(* IEC 61131-3 sources: SortJet_MasterSPS_Aufbau.fbsproj/08_POUs/Basis Programmbausteine, 6 files *)

(* ---- AutomatischeFachaufnahme.prg.st ---- *)
(* METADATA
{
	"v3Meta": {
		"objectGuid": "2dd67d59-9d65-422a-a9a5-a54784296135"
	}
}
*)
PROGRAM AutomatischeFachaufnahme
VAR_INPUT

  // BOOLEAN
  bpStarteFachaufnahme : BOOL := FALSE;
  bpAktiv              : BOOL := TRUE;

  // WORD
  wpMMINummer  : WORD;

  // POINTER
  ptQuerfahrtShuttle : REFERENCE TO Rexroth_ctrlX_Drive_Eckelmann_MC_V01_02_02;

  // REF
  Shuttle : REFERENCE TO Shuttle_FB_V01_00_00;

END_VAR

VAR

  // STEP
  steplAufnahme            : STEPS_TE;

  // WORD

  // REAL
  rlLetztePosition         : REAL;
  rlMerkerGeschwindigkeit  : real;

  // POINTER
  ptlAnalogwertChannel1  : REFERENCE TO INT;
  ptlAnalogwertChannel2  : REFERENCE TO INT;

END_VAR

VAR CONSTANT

  // WORD
  wGeschwindigkeitFachaufnahme : WORD := 5;
  wDefaultHandgeschwindigkeit  : WORD := 300;

END_VAR

//-------------------------------------------------------------------------------------------------
// AUTOMATISIERTE FACHAUFNAHME
//-------------------------------------------------------------------------------------------------
(* Anmerkung:
   - Shuttle-Koordinationsbaustein zur Fachaufnahme
*)
IF ( bpAktiv ) THEN

  (* Hinweis:
     - Starten der Fachaufnahme
  *)
  Shuttle REF= aShuttle[wpMMINummer];
  IF NOT __ISVALIDREF(Shuttle) THEN
    RETURN;
  ELSE
    ptQuerfahrtShuttle    REF= Shuttle.Querfahrt.Antrieb;
    ptlAnalogwertChannel1 REF= Shuttle.in_iAnalogwertChannel1;
    ptlAnalogwertChannel2 REF= Shuttle.in_iAnalogwertChannel2;
  END_IF

  (* Hinweis:
     - Starten der Fachaufnahme
  *)
  IF ( bpStarteFachaufnahme ) THEN

    IF ( __ISVALIDREF(ptQuerfahrtShuttle) ) THEN

      CASE steplAufnahme OF

        // -----------------------------------------------------------------------
        STEP_0_E:
          rlMerkerGeschwindigkeit :=  ptQuerfahrtShuttle.ppAntriebsInformationen.rpHandGeschwindigkeit;
          ptQuerfahrtShuttle.ppAntriebsInformationen.rpHandGeschwindigkeit := wGeschwindigkeitFachaufnahme;

          steplAufnahme:= STEP_10_E;

        // -----------------------------------------------------------------------
        STEP_10_E:
          IF (  ( ptQuerfahrtShuttle.rpIstPosition <> rlLetztePosition )
               AND ( ptQuerfahrtShuttle.rpIstPosition <> 0 ) )
          THEN

            rlLetztePosition := ptQuerfahrtShuttle.rpIstPosition;

            (* Hinweis:
               - Nachricht an das HMI
            *)
            rSPS2MMIFachaufnahmePosition   := rlLetztePosition;
            wSPS2MMIFachaufnahmeAnalogwert := TO_WORD(ptlAnalogwertChannel1);
            MsgToMmi( SB0_SPS_FACHAUFNAHMEDATEN );
          END_IF

      END_CASE

    ELSE
      ;

    END_IF

  END_IF

  IF ( NOT bpStarteFachaufnahme ) THEN

    IF ( steplAufnahme > STEP_0_E ) THEN
      steplAufnahme := STEP_0_E;
      ptQuerfahrtShuttle.ppAntriebsInformationen.rpHandGeschwindigkeit := SEL( rlMerkerGeschwindigkeit <> 0, wDefaultHandgeschwindigkeit, rlMerkerGeschwindigkeit ) ;
      rlMerkerGeschwindigkeit := 0;
    END_IF

  END_IF

END_IF
END_PROGRAM

(* ---- CheckReset.prg.st ---- *)
(* METADATA
{
	"v3Meta": {
		"objectGuid": "ed448837-b746-4b1a-b2e7-236797e04e0f"
	}
}
*)
PROGRAM CheckReset
VAR
  wlIndexAutomatikkreis,
  wlIndexStation : WORD;
END_VAR

FOR wlIndexAutomatikkreis := cERSTER_AUTOMATIKKREIS TO cLETZTER_AUTOMATIKKREIS DO

  agbResetAktiv[wlIndexAutomatikkreis] := FALSE;

  FOR wlIndexStation := cERSTE_STATION TO cLETZTE_STATION DO
    IF starrStationBasisParameter[wlIndexStation].bReset AND_THEN StationInAutomatikkreis(starrStationBasisParameter[wlIndexStation].stMKs.eaAutomatikkreis, wlIndexAutomatikkreis) THEN
      agbResetAktiv[wlIndexAutomatikkreis] := TRUE;
      EXIT;
    END_IF
  END_FOR

  // Schleife des AK eine Iteration weiter
  IF agbResetAktiv[wlIndexAutomatikkreis] THEN
    CONTINUE;
  END_IF

  FOR wlIndexStation := cERSTES_SHUTTLE TO cLETZTES_SHUTTLE DO
    IF starrShuttleBasisParameter[wlIndexStation].bReset AND_THEN StationInAutomatikkreis(starrShuttleBasisParameter[wlIndexStation].stMKs.eaAutomatikkreis, wlIndexAutomatikkreis) THEN
      agbResetAktiv[wlIndexAutomatikkreis] := TRUE;
      EXIT;
    END_IF
  END_FOR

  // Schleife des AK eine Iteration weiter
  IF agbResetAktiv[wlIndexAutomatikkreis] THEN
    CONTINUE;
  END_IF

  FOR wlIndexStation := cERSTES_TRANSFERSHUTTLE TO cLETZTES_TRANSFERSHUTTLE DO
    IF starrTransferShuttleBasisParameter[wlIndexStation].bReset AND_THEN StationInAutomatikkreis(starrTransferShuttleBasisParameter[wlIndexStation].stMKs.eaAutomatikkreis, wlIndexAutomatikkreis) THEN
      agbResetAktiv[wlIndexAutomatikkreis] := TRUE;
      EXIT;
    END_IF
  END_FOR

  // Schleife des AK eine Iteration weiter
  IF agbResetAktiv[wlIndexAutomatikkreis] THEN
    CONTINUE;
  END_IF

  FOR wlIndexStation := cERSTE_FAECHERWAGENSTATIONS_NR TO cLETZTE_FAECHERWAGENSTATIONS_NR DO
    IF starrFaecherwagenBasisParameter[wlIndexStation].bReset AND_THEN StationInAutomatikkreis(starrFaecherwagenBasisParameter[wlIndexStation].stMKs.eaAutomatikkreis, wlIndexAutomatikkreis) THEN
      agbResetAktiv[wlIndexAutomatikkreis] := TRUE;
      EXIT;
    END_IF
  END_FOR

  // Schleife des AK eine Iteration weiter
  IF agbResetAktiv[wlIndexAutomatikkreis] THEN
    CONTINUE;
  END_IF

  FOR wlIndexStation := cERSTE_FREMDANLAGE_EINLAUF TO cLETZTE_FREMDANLAGE_EINLAUF DO
    IF starrFremdanlageEinlaufStationBasisParameter[wlIndexStation].bReset AND_THEN StationInAutomatikkreis(starrFremdanlageEinlaufStationBasisParameter[wlIndexStation].stMKs.eaAutomatikkreis, wlIndexAutomatikkreis) THEN
      agbResetAktiv[wlIndexAutomatikkreis] := TRUE;
      EXIT;
    END_IF
  END_FOR

  // Schleife des AK eine Iteration weiter
  IF agbResetAktiv[wlIndexAutomatikkreis] THEN
    CONTINUE;
  END_IF

  FOR wlIndexStation := cERSTE_FREMDANLAGE_AUSLAUF TO cLETZTE_FREMDANLAGE_AUSLAUF DO
    IF starrFremdanlageAuslaufStationBasisParameter[wlIndexStation].bReset AND_THEN StationInAutomatikkreis(starrFremdanlageAuslaufStationBasisParameter[wlIndexStation].stMKs.eaAutomatikkreis, wlIndexAutomatikkreis) THEN
      agbResetAktiv[wlIndexAutomatikkreis] := TRUE;
      EXIT;
    END_IF
  END_FOR

END_FOR
END_PROGRAM

(* ---- ErsteUndLetzteScheibeBits.prg.st ---- *)
(* METADATA
{
	"v3Meta": {
		"objectGuid": "2dfa9b46-65fe-42f1-b72f-b251bddaa00a"
	}
}
*)
PROGRAM ErsteUndLetzteScheibeBits
VAR_INPUT

  // WORD
  wpErsteUndLetzteScheibe : WORD;

END_VAR
VAR_OUTPUT

  // WORD
  wpLetzteScheibe,
  wpErsteScheibe   : WORD;

END_VAR
VAR

  // WORD
  wlMerkerErsteUndLetzteScheibe  : WORD;

END_VAR
VAR CONSTANT

  // WORD
  cBIT_MASKE_LETZTE_SCHEIBE  : WORD := 2#0000000011111111;

END_VAR

//-------------------------------------------------------------------------------------------------
// BAUSTEIN: LOGIK
//-------------------------------------------------------------------------------------------------

(* Hinweis:
   - Erste Scheibe
*)
wlMerkerErsteUndLetzteScheibe := wpErsteUndLetzteScheibe;
wpLetzteScheibe := wlMerkerErsteUndLetzteScheibe AND cBIT_MASKE_LETZTE_SCHEIBE;

(* Hinweis:
   - Letzte Scheibe
*)
wlMerkerErsteUndLetzteScheibe := wpErsteUndLetzteScheibe;
wpErsteScheibe := SHR(wlMerkerErsteUndLetzteScheibe, 8);
END_PROGRAM

(* ---- Schrittketten_Logger.prg.st ---- *)
(* METADATA
{
	"v3Meta": {
		"objectGuid": "cb3b1eb5-1dc3-4d16-abd2-ade96f8e42d9"
	}
}
*)
PROGRAM Schrittketten_Logger
VAR

  // WORD
  i              : WORD;
  j              : WORD;
  wiSchrittkette : ARRAY[0..7] OF WORD;
  wlSchrittkette : ARRAY[0..7,0..31] OF WORD;

  // STRING
  sBezeichnung   : ARRAY[0..7] OF STRING;

END_VAR
sBezeichnung[0]   := ' - ';
wiSchrittkette[0] := 0;

sBezeichnung[1]   := ' - ';
wiSchrittkette[1] := 0;

sBezeichnung[2]   :=  ' - ';
wiSchrittkette[2] :=  0;

sBezeichnung[3]   :=  ' - ';
wiSchrittkette[3] :=  0;

sBezeichnung[4]   := ' - ';
wiSchrittkette[4] := 0;

sBezeichnung[5]   := ' - ';
wiSchrittkette[5] := 0;

sBezeichnung[6]   := ' - ';
wiSchrittkette[6] := 0;

sBezeichnung[7]   := ' - ';
wiSchrittkette[7] := 0;

FOR i := 0 TO 7 DO

  IF(wiSchrittkette[i] <> wlSchrittkette[i,31])THEN;

    FOR j := 0 TO 30 DO
      wlSchrittkette[i,j] := wlSchrittkette[i,j+1];
    END_FOR

    wlSchrittkette[i,31] := wiSchrittkette[i];
  END_IF

END_FOR
END_PROGRAM

(* ---- StartUpCheck.prg.st ---- *)
(* METADATA
{
	"v3Meta": {
		"objectGuid": "11193127-30f6-42cb-ab25-4fe444daee5f"
	}
}
*)
PROGRAM StartUpCheck
VAR
  aUsedAchsIDs : ARRAY [0..65] OF BOOL;
  aUsedMeldungsnummern : ARRAY [0..2500] OF BOOL;
  aUsedStationNrIntern : ARRAY [cERSTES_SHUTTLE..cLETZTE_FREMDANLAGE_EINLAUF] OF BOOL;
  aUsedStationNrSPS    : ARRAY [cERSTES_SHUTTLE..cLETZTE_FREMDANLAGE_EINLAUF] OF BOOL;

  i : WORD;
  k : WORD;
  cLOG_HANDLE : RTS_IEC_HANDLE := RTS_INVALID_HANDLE;
  NullRef : REFERENCE TO BOOL;
END_VAR

FOR i := cERSTES_SHUTTLE TO cLETZTES_SHUTTLE DO
  // wAchsID in den Antriebsinformationen prüfen - niccht doppelt vergeben
  FOR k := cWAND_1 TO cANZAHL_WAENDE DO
    CheckAchsID(starrShuttleBasisParameter[i].stAntriebsparameter.stGlastransport[k].wAchsID);
    CheckAchsID(starrShuttleBasisParameter[i].stAntriebsparameter.stGlastransportSlave[k].wAchsID);
    CheckAchsID(starrShuttleBasisParameter[i].stAntriebsparameter.stWandverstellung[k].wAchsID);
  END_FOR
  CheckAchsID(starrShuttleBasisParameter[i].stAntriebsparameter.stDrehen.wAchsID);
  CheckAchsID(starrShuttleBasisParameter[i].stAntriebsparameter.stKippen.wAchsID);
  CheckAchsID(starrShuttleBasisParameter[i].stAntriebsparameter.stMessachse.wAchsID);
  CheckAchsID(starrShuttleBasisParameter[i].stAntriebsparameter.stQuerfahrt.wAchsID);
  // Konfigurierete Automatikkreise prüfen
  CheckAutomatikkreis(starrShuttleBasisParameter[i]);
  // Konfiguriereten StationsTyp prüfen
  CheckStationsTyp(starrShuttleBasisParameter[i]);
  // Konfigurierete Meldungsnummer prüfen
  CheckMeldungsnummer(starrShuttleBasisParameter[i]);
  // Konfigurierete Stationsnummern prüfen
  CheckStationsnummern(starrShuttleBasisParameter[i]);
  // Konfigurierte Lage der letzten Scheibe prüfen
  checkGlastransportOptionen(starrShuttleBasisParameter[i], TRUE);
END_FOR

FOR i := cERSTES_TRANSFERSHUTTLE TO cLETZTES_TRANSFERSHUTTLE DO
  FOR k := cWAND_1 TO cANZAHL_WAENDE DO
    CheckAchsID(starrTransfershuttleBasisParameter[i].stAntriebsparameter.stGlastransport[k].wAchsID);
    CheckAchsID(starrTransfershuttleBasisParameter[i].stAntriebsparameter.stGlastransportSlave[k].wAchsID);
    CheckAchsID(starrTransfershuttleBasisParameter[i].stAntriebsparameter.stWandverstellung[k].wAchsID);
  END_FOR
  CheckAchsID(starrTransfershuttleBasisParameter[i].stAntriebsparameter.stDrehen.wAchsID);
  CheckAchsID(starrTransfershuttleBasisParameter[i].stAntriebsparameter.stKippen.wAchsID);
  CheckAchsID(starrTransfershuttleBasisParameter[i].stAntriebsparameter.stMessachse.wAchsID);
  CheckAchsID(starrTransfershuttleBasisParameter[i].stAntriebsparameter.stQuerfahrt.wAchsID);
  // Konfigurierete Automatikkreise prüfen
  CheckAutomatikkreis(starrTransfershuttleBasisParameter[i]);
  // Konfiguriereten StationsTyp prüfen
  CheckStationsTyp(starrTransfershuttleBasisParameter[i]);
  // Konfigurierete Meldungsnummer prüfen
  CheckMeldungsnummer(starrTransfershuttleBasisParameter[i]);
  // Konfigurierete Stationsnummern prüfen
  CheckStationsnummern(starrTransfershuttleBasisParameter[i]);
END_FOR

FOR i := cERSTE_STATION TO cLETZTE_STATION DO
  FOR k := cWAND_1 TO cANZAHL_WAENDE DO
    CheckAchsID(starrStationBasisParameter[i].stAntriebsparameter.stGlastransport[k].wAchsID);
    CheckAchsID(starrStationBasisParameter[i].stAntriebsparameter.stGlastransportSlave[k].wAchsID);
    IF __ISVALIDREF(starrStationBasisParameter[i].stAntriebsparameter.stGlastransportY) THEN
      CheckAchsID(starrStationBasisParameter[i].stAntriebsparameter.stGlastransportY[k].wAchsID);
    END_IF
    IF __ISVALIDREF(starrStationBasisParameter[i].stAntriebsparameter.stGlastransportYSlave) THEN
      CheckAchsID(starrStationBasisParameter[i].stAntriebsparameter.stGlastransportYSlave[k].wAchsID);
    END_IF
    CheckAchsID(starrStationBasisParameter[i].stAntriebsparameter.stWandverstellung[k].wAchsID);
  END_FOR
  CheckAchsID(starrStationBasisParameter[i].stAntriebsparameter.stDrehen.wAchsID);
  CheckAchsID(starrStationBasisParameter[i].stAntriebsparameter.stKippen.wAchsID);
  CheckAchsID(starrStationBasisParameter[i].stAntriebsparameter.stMessachse.wAchsID);
  CheckAchsID(starrStationBasisParameter[i].stAntriebsparameter.stQuerfahrt.wAchsID);
  // Konfigurierete Automatikkreise prüfen
  CheckAutomatikkreis(starrStationBasisParameter[i]);
  // Konfiguriereten StationsTyp prüfen
  CheckStationsTyp(starrStationBasisParameter[i]);
  // Konfigurierete Meldungsnummer prüfen
  CheckMeldungsnummer(starrStationBasisParameter[i]);
  // Konfigurierete Stationsnummern prüfen
  CheckStationsnummern(starrStationBasisParameter[i]);
  // Konfigurierte Lage der letzten Scheibe prüfen
  checkGlastransportOptionen(starrStationBasisParameter[i], FALSE);
END_FOR

checkMKVerfahrparameter();
checkZentralschmierung();
checkAutomatikkreiseMK();
checkSicherheitskreiseMK();
checkDurchgaenge();
END_PROGRAM

(* ---- VailiderenTransfershuttleVerbund.prg.st ---- *)
(* METADATA
{
	"v3Meta": {
		"objectGuid": "53cd760f-4cde-42f5-90aa-7a00051f7bed"
	}
}
*)
PROGRAM VailiderenTransfershuttleVerbund
VAR
END_VAR

VAR_INPUT

  // WORD
  wTransferstation1 : WORD;
  wTransferstation2 : WORD;

END_VAR

VAR_OUTPUT

  // BOOL
  bpFehler : BOOL;

  // WORD
  wTransferstationMaster : WORD;
  wTransferstationSlave  : WORD;

END_VAR

//-------------------------------------------------------------------------------------------------
// BAUSTEIN: LOGIK
//-------------------------------------------------------------------------------------------------
(* Hinweis:
   - Fehler ggf. zuruecksetzen
*)
bpFehler := FALSE;

(* Hinweis:
   - Validieren
*)
IF (  ( PruefungWertImIntervall(wTransferstation1, cERSTES_TRANSFERSHUTTLE , cLETZTES_TRANSFERSHUTTLE ) )
     AND ( PruefungWertImIntervall(wTransferstation2, cERSTES_TRANSFERSHUTTLE , cLETZTES_TRANSFERSHUTTLE ) ) )
THEN

  IF (      ( starrTransfershuttleBasisParameter[wTransferstation1].stMKs.stStationsOptionen.stTransfershuttle.bMasterStation = TRUE )
       AND NOT ( starrTransfershuttleBasisParameter[wTransferstation2].stMKs.stStationsOptionen.stTransfershuttle.bMasterStation = TRUE ) )
  THEN
    wTransferstationMaster := wTransferstation1;
    wTransferstationSlave  := wTransferstation2;

  ELSIF (   ( starrTransfershuttleBasisParameter[wTransferstation2].stMKs.stStationsOptionen.stTransfershuttle.bMasterStation = TRUE )
          AND NOT ( starrTransfershuttleBasisParameter[wTransferstation1].stMKs.stStationsOptionen.stTransfershuttle.bMasterStation = TRUE ) )
  THEN
    wTransferstationMaster := wTransferstation2;
    wTransferstationSlave  := wTransferstation1;

  ELSE
    bpFehler := TRUE;

    wTransferstationMaster := wTransferstation1;
    wTransferstationSlave  := wTransferstation2;

    wpgFehlerdaten[0] := wTransferstation1;
    wpgFehlerdaten[0] := wTransferstation2;
    SpsHinweis( eFehler_Station,
                cMELDUNG_TS_KONNTE_KEIN_MASTER_TS_ERMITTELT_WERDEN,
                wTransferstation1,
                AutomatikkreisBestimmen(starrTransfershuttleBasisParameter[wTransferstation1].stMKs.stStationsNummern.NummerSPS),
                wpgFehlerdaten );

  (* Anmerkung:
     - Hier muesste ein fehler geworfen werden
  *)

  END_IF

ELSE
  bpFehler := TRUE;

(* Anmerkung:
   - Hier muesste ein fehler geworfen werden
*)

END_IF
END_PROGRAM
